// TIA Portal V21 program export: 0 tag tables, 0 data types, 0 data blocks, 2 code blocks (in call order from the OBs), 0 instance data blocks

ORGANIZATION_BLOCK "Edges"   // OB1, LAD
   VAR_TEMP   // added for the SCL form of the ladder/FBD networks
      _w1 : Bool;
   END_VAR
BEGIN

REGION Network 1: Rising edge
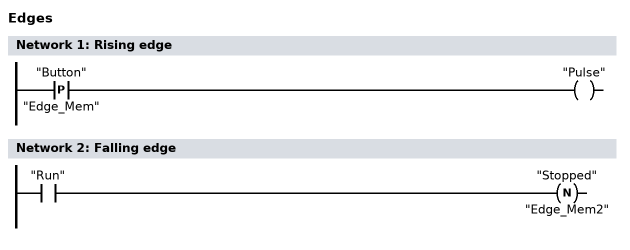
   #_w1 := "Button" AND NOT "Edge_Mem";   // rising edge of "Button"
   "Edge_Mem" := "Button";
   "Pulse" := #_w1;
END_REGION

REGION Network 2: Falling edge
   "Stopped" := NOT "Run" AND "Edge_Mem2";   // falling edge
   "Edge_Mem2" := "Run";
END_REGION
END_ORGANIZATION_BLOCK

FUNCTION_BLOCK "Mixed"   // FB1, LAD
BEGIN

REGION Network 1: Unknown part
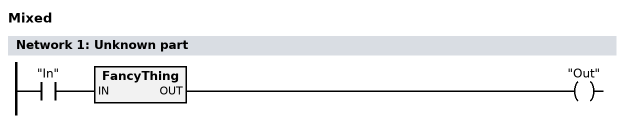
   // no SCL statement known for FancyThing: written as a call
   "Out" := FancyThing("In");
END_REGION

REGION Network 2 (SCL): SCL inside
END_REGION

REGION Network 3: Empty
END_REGION
END_FUNCTION_BLOCK
